Fanuc KAREL source: KO00033.KL

PROGRAM KO00033
%NOLOCKGROUP
%ENVIRONMENT MIR
VAR
  P1: POSITION
  P2: POSITION
  F: BOOLEAN
  OUT: POSITION
BEGIN
  F = TRUE
  OUT = MIRROR(P1, P2, F)
END KO00033
